(* Processor test double that counts what the simple processor does with each span. *)
FUNCTION_BLOCK FB_SpanProcessor_ForInspection EXTENDS FB_SpanProcessor_Simple
VAR_OUTPUT
	enrichedCount: UDINT;
	exportedCount: UDINT;
	tickCount: UDINT;
	enrichedBeforeExport: BOOL;
	lastSpanName: T_MaxString;
END_VAR

METHOD enrich
VAR_IN_OUT
	span: FB_Span;
END_VAR
THIS^.enrichedCount := THIS^.enrichedCount + 1;
END_METHOD

METHOD export
VAR_INPUT
	span: REFERENCE TO FB_Span;
END_VAR
THIS^.exportedCount := THIS^.exportedCount + 1;
THIS^.enrichedBeforeExport := THIS^.enrichedCount = THIS^.exportedCount;
IF span.name <> 0 AND_THEN span.name^.pString <> 0 THEN
	THIS^.lastSpanName := span.name^.pString^;
END_IF
END_METHOD

METHOD tick
THIS^.tickCount := THIS^.tickCount + 1;
END_METHOD

END_FUNCTION_BLOCK

(* stored: Version 1.1.0.1
   POU FB_SpanProcessor_ForInspection: Id {eb9c9fd4-ddec-40c9-a62f-4563a975c8c6}, SpecialFunc None
   Method enrich: Id {fded2ebe-3674-4697-8816-96388bc115de}
   Method export: Id {51792d96-aa8f-4ed6-afbe-c57e4fc200b9}
   Method tick: Id {ad98e666-c3e3-4518-9182-8b730792294b} *)
